(* PLC project Vn_ton_boxes_on_pins, Beckhoff Automation GmbH TwinCAT PLC Control 3.5.13.21 *)
(* stored: creationDateTime 1970-01-01T00:00:00 *)

PROGRAM Vn_ton_boxes_on_pins

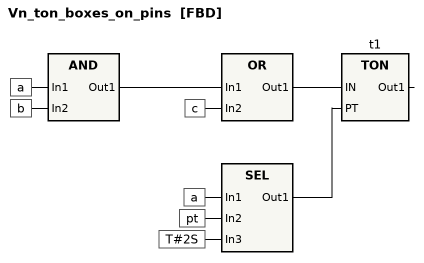
(* FBD diagram, written out as Structured Text *)
t1(IN := a AND b OR c, PT := SEL(a, pt, T#2S));
END_PROGRAM
